FUNCTION_BLOCK Preparador_Vibropac_HMI (* Service Interface Function Block Type *)
  (* Standard: 61499-2 *)
  (* Version 1.0, 19/10/2026, Hidryco, Hidryco, IHM do Preparador_Vibropac *)
  PACKAGE Hidryco.HidrycoLib;
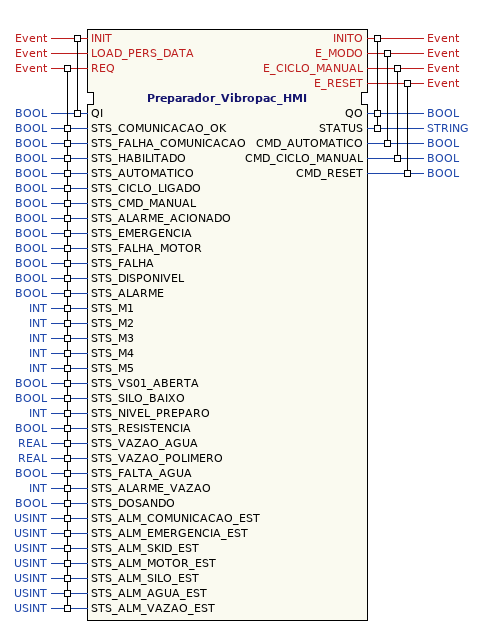
  EVENT_INPUT
    INIT WITH QI;
    LOAD_PERS_DATA; (* Reenvia os parametros persistentes *)
    REQ WITH STS_COMUNICACAO_OK, STS_FALHA_COMUNICACAO, STS_HABILITADO, STS_AUTOMATICO, STS_CICLO_LIGADO, STS_CMD_MANUAL, STS_ALARME_ACIONADO, STS_EMERGENCIA, STS_FALHA_MOTOR, STS_FALHA, STS_DISPONIVEL, STS_ALARME, STS_M1, STS_M2, STS_M3, STS_M4, STS_M5, STS_VS01_ABERTA, STS_SILO_BAIXO, STS_NIVEL_PREPARO, STS_RESISTENCIA, STS_VAZAO_AGUA, STS_VAZAO_POLIMERO, STS_FALTA_AGUA, STS_ALARME_VAZAO, STS_DOSANDO, STS_ALM_COMUNICACAO_EST, STS_ALM_EMERGENCIA_EST, STS_ALM_SKID_EST, STS_ALM_MOTOR_EST, STS_ALM_SILO_EST, STS_ALM_AGUA_EST, STS_ALM_VAZAO_EST; (* Atualizacao de status *)
  END_EVENT
  EVENT_OUTPUT
    INITO WITH QO, STATUS;
    E_MODO WITH CMD_AUTOMATICO;
    E_CICLO_MANUAL WITH CMD_CICLO_MANUAL;
    E_RESET WITH CMD_RESET;
  END_EVENT
  VAR_INPUT
    QI : BOOL;
    STS_COMUNICACAO_OK : BOOL; (* Comunicacao Modbus com o CLP do skid OK *)
    STS_FALHA_COMUNICACAO : BOOL; (* Falha de comunicacao com o CLP do skid *)
    STS_HABILITADO : BOOL; (* Instancia habilitada (FALSE = equipamento futuro) *)
    STS_AUTOMATICO : BOOL; (* Ciclo comandado pelo processo (automatico) *)
    STS_CICLO_LIGADO : BOOL; (* Comando de ciclo remoto ligado (4001 = 1) *)
    STS_CMD_MANUAL : BOOL; (* Comando manual de ciclo (modo manual) *)
    STS_ALARME_ACIONADO : BOOL; (* Alarme acionado no skid (4005) *)
    STS_EMERGENCIA : BOOL; (* Botao de emergencia do skid acionado (4006) *)
    STS_FALHA_MOTOR : BOOL; (* Algum motor do skid em falha *)
    STS_FALHA : BOOL; (* Skid em falha (alarme, emergencia ou motor) *)
    STS_DISPONIVEL : BOOL; (* Pode ser ligado pelo automatico agora *)
    STS_ALARME : BOOL; (* Algum alarme do skid *)
    STS_M1 : INT; (* Status M1 agitador do tanque de mistura (4007): 0 parado, 1 funcionando, 2 falha *)
    STS_M2 : INT; (* Status M2 agitador do tanque de maturacao (4008): 0 parado, 1 funcionando, 2 falha *)
    STS_M3 : INT; (* Status M3 dosador volumetrico (4009): 0 parado, 1 funcionando, 2 falha *)
    STS_M4 : INT; (* Status M4 bomba dosadora M4 (4010): 0 parado, 1 funcionando, 2 falha *)
    STS_M5 : INT; (* Status M5 bomba dosadora M5 (4011): 0 parado, 1 funcionando, 2 falha *)
    STS_VS01_ABERTA : BOOL; (* Solenoide de agua VS-01 aberta (4012) *)
    STS_SILO_BAIXO : BOOL; (* Silo de polimero em po com nivel baixo LSL-01 (4013 = 0) *)
    STS_NIVEL_PREPARO : INT; (* Nivel LS1: 0 muito baixo, 1 baixo, 2 alto, 3 muito alto (4014) *)
    STS_RESISTENCIA : BOOL; (* Resistencia de aquecimento RA-01 ligada (4015) *)
    STS_VAZAO_AGUA : REAL; (* Vazao de agua FIT-01 (%) (4016, 0-1000) *)
    STS_VAZAO_POLIMERO : REAL; (* Vazao de polimero preparado FIT-02 (%) (4017, 0-1000) *)
    STS_FALTA_AGUA : BOOL; (* Alarme de falta d agua (4018) *)
    STS_ALARME_VAZAO : INT; (* Alarme de vazao de polimero: 0 sem, 1 baixa, 2 alta (4019) *)
    STS_DOSANDO : BOOL; (* Bomba dosadora M4 ou M5 funcionando *)
    STS_ALM_COMUNICACAO_EST : USINT; (* Estado do ALARM_BIT (0 normal, 1 ativo reconhecido, 2 ativo nao reconhecido, 3 saiu nao reconhecido, 4 ativo e saiu nao reconhecido) *)
    STS_ALM_EMERGENCIA_EST : USINT; (* Estado do ALARM_BIT (0 normal, 1 ativo reconhecido, 2 ativo nao reconhecido, 3 saiu nao reconhecido, 4 ativo e saiu nao reconhecido) *)
    STS_ALM_SKID_EST : USINT; (* Estado do ALARM_BIT (0 normal, 1 ativo reconhecido, 2 ativo nao reconhecido, 3 saiu nao reconhecido, 4 ativo e saiu nao reconhecido) *)
    STS_ALM_MOTOR_EST : USINT; (* Estado do ALARM_BIT (0 normal, 1 ativo reconhecido, 2 ativo nao reconhecido, 3 saiu nao reconhecido, 4 ativo e saiu nao reconhecido) *)
    STS_ALM_SILO_EST : USINT; (* Estado do ALARM_BIT (0 normal, 1 ativo reconhecido, 2 ativo nao reconhecido, 3 saiu nao reconhecido, 4 ativo e saiu nao reconhecido) *)
    STS_ALM_AGUA_EST : USINT; (* Estado do ALARM_BIT (0 normal, 1 ativo reconhecido, 2 ativo nao reconhecido, 3 saiu nao reconhecido, 4 ativo e saiu nao reconhecido) *)
    STS_ALM_VAZAO_EST : USINT; (* Estado do ALARM_BIT (0 normal, 1 ativo reconhecido, 2 ativo nao reconhecido, 3 saiu nao reconhecido, 4 ativo e saiu nao reconhecido) *)
  END_VAR
  VAR_OUTPUT
    QO : BOOL; (* Event Output Qualifier *)
    STATUS : STRING; (* Service Status *)
    CMD_AUTOMATICO : BOOL; (* TRUE = automatico (ciclo pelo processo); persistente *)
    CMD_CICLO_MANUAL : BOOL; (* Manual: TRUE liga o ciclo remoto *)
    CMD_RESET : BOOL; (* Reset do skid (4002) e reconhecimento dos alarmes *)
  END_VAR
  SERVICE /
    SEQUENCE 
    END_SEQUENCE
  END_SERVICE
END_FUNCTION_BLOCK
